Fanuc KAREL source: KA00140.KL

PROGRAM KA00140
%NOLOCKGROUP
VAR
  SRC: ARRAY[2] OF SHORT
  DST: JOINTPOS
BEGIN
  SRC[1] = 2
  DST = SRC[1]
END KA00140
